// Generated by voz_llm_plc_agent
// Target: Siemens TIA Portal V18 - SCL external source
// Review and compile before any download to physical hardware.

FUNCTION_BLOCK "PLC_PRG"
{ S7_Optimized_Access := 'TRUE' }
VERSION : 0.1
VAR_INPUT
   I_Maintenance_Mode : Bool := FALSE;
   I_Start : Bool := FALSE;
   I_Emergency : Bool := FALSE;
   I_Maintenance : Bool := FALSE;
END_VAR
VAR_OUTPUT
   Q_Motor_Enable : Bool := FALSE;
END_VAR
BEGIN
(* Bloqueo de arranque durante mantenimiento *)
IF #I_Maintenance_Mode THEN
    #Q_Motor_Enable := FALSE;
ELSE
    #Q_Motor_Enable := #I_Start AND NOT #I_Emergency;
END_IF;
END_FUNCTION_BLOCK

DATA_BLOCK "DB_PLC_PRG"
{ S7_Optimized_Access := 'TRUE' }
VERSION : 0.1
NON_RETAIN
"PLC_PRG"
BEGIN
END_DATA_BLOCK

ORGANIZATION_BLOCK "Main"
{ S7_Optimized_Access := 'TRUE' }
VERSION : 0.1
BEGIN
   "DB_PLC_PRG"(
      I_Maintenance_Mode := "I_Maintenance_Mode",
      I_Start := "I_Start",
      I_Emergency := "I_Emergency",
      Q_Motor_Enable => "Q_Motor_Enable",
      I_Maintenance := "I_Maintenance"
   );
END_ORGANIZATION_BLOCK
